(* CODESYS project stringhandler.library
   Company: KOSTAL GmbH & Co.KG
   Version: 2019.3.4.0
   DefaultNamespace: KOSTAL.TC3.Components.Stringhandler
   Title: KOSTAL.TC3.Components.Stringhandler
   Placeholder: KOSTAL.TC3.Components.Stringhandler
   Author: Frank Dümpelmann
   DocFormat: reStructuredText

Project tree, tasks and I/O mapping:
  libraries: KOSTAL.TC3.Components.listOfString, 2019.2.2.0 (KOSTAL GmbH & Co.KG); KOSTAL.TC3.Core.functionResponse, 2019.0.3.0 (KOSTAL GmbH & Co.KG); KOSTAL.TC3.Core.Settings, 2019.0.1.0 (KOSTAL GmbH & Co.KG); Tc2_Math, 3.3.1.0 (Beckhoff Automation GmbH); Tc2_Standard, 3.3.3.0 (Beckhoff Automation GmbH); Tc2_System, 3.4.26.0 (Beckhoff Automation GmbH); Tc2_Utilities, 3.3.54.0 (Beckhoff Automation GmbH); Tc3_Module, 3.3.21.0 (Beckhoff Automation GmbH)
  DUT/
    data type E_ALIGNMENT
  POU/
    obsolete/
      function F_CONCAT [ST]
      function F_Format [ST]
      function F_Text_Clear [ST]
      function block FB_Split [ST]: _pResult_clear, _settingsControl, Delimiter, pResults, sizeOfResultArray, split, status
    function F_FLOAT_TO_STRING [ST]
    function F_FormatMask [ST]
    function F_FormatNoMask [ST]
    function F_LCASE [ST]
    function F_LREAL_TO_STRING [ST]
    function F_REAL_TO_STRING [ST]
    function F_Replace [ST]
    function F_UCASE [ST]
    function block FB_CONCAT [ST]: addContent, clear, FB_exit, getResult, new
    function block FB_SplitEx [ST]: _settingsControl, clear, Delimiter, FB_exit, FB_init, getElement, maxElement, setElement, split, status
    function block FB_UrlEscape [ST]: Execute
  Project Information/
    function F_GetCompany [ST]
    function F_GetTitle [ST]
    function F_GetVersion [ST]
  Version/
    global variables Global_Version
  global variables GVL_CONSTANT
*)

// DUT/E_ALIGNMENT
TYPE E_ALIGNMENT :
	(
		LEFT 	:= 0,
		RIGHT	:= 1,
		CENTER	:= 2
	);
END_TYPE

// Version/Global_Version
{attribute 'TcGenerated'}
{attribute 'no-analysis'}
{attribute 'linkalways'}
// This function has been automatically generated from the project information.
VAR_GLOBAL CONSTANT
	{attribute 'const_non_replaced'}
	stLibVersion_KOSTAL_TC3_Components_Stringhandler : ST_LibVersion := (iMajor := 2019, iMinor := 3, iBuild := 4, iRevision := 0, nFlags := 1, sVersion := '2019.3.4.0');
END_VAR

// GVL_CONSTANT
{attribute 'qualified_only'}
VAR_GLOBAL CONSTANT
	
(*
65 A 	97 a 
66 B 	98 b 
67 C 	99 c 
68 D 	100 d 
69 E 	101 e 
70 F 	102 f 
71 G 	103 g 
72 H 	104 h 
73 I 	105 i 
74 J 	106 j 
75 K 	107 k 
76 L 	108 l 
77 M 	109 m 
78 N 	110 n 
79 O 	111 o 
80 P 	112 p 
81 Q 	113 q 
82 R 	114 r 
83 S 	115 s 
84 T 	116 t 
85 U 	117 u 
86 V 	118 v 
87 W 	119 w 
88 X 	120 x 
89 Y 	121 y 
90 Z 	122 z
*)

	START_UCASE	: BYTE:= 65;	//BYTE:= 65
	END_UCASE		: BYTE:= 90;	//BYTE:= 90
	START_LCASE	: BYTE:= 97;	//BYTE:= 97
	END_LCASE		: BYTE:= 122;	//BYTE:= 122
	OFFSET			: BYTE:= 32;	//BYTE:= 32

	OVERFLOW	: STRING:= 'OVERFLOW';
	
END_VAR

// POU/obsolete/F_CONCAT
(*

:Author: Frank Dümpelmann <f.duempelmann@kostal.com>, Martin Hundt <m.hundt@kostal.com>
:Date: 2018-10-29

Function
========
Concatination of variable number of lines to one line with maximum 255 chars

Usage notes
===============
Won't work with arrays shorter than 255 chars

Parameters
======================
| P_Line_1		: POINTER TO STRING(255) - Pointer to first element of an array[1..numberOfLines] OF STRING(255)
| numberOfLines	: USINT - defines the number of elements of the Array 

Return Value
============
String(255) - Concatination of the array's elements

Usage sample:
=============

.. code:: 

	PROGRAM MAIN
	VAR
		_aStrings	: ARRAY [0..4] OF STRING(255);
		_output 	: STRING(255); 
	END_VAR
	
	_aStrings[0] := 'Kostal';
	_aStrings[1] := ' ';
	_aStrings[2] := 'Automobil';
	_aStrings[3] := ' ';
	_aStrings[4] := 'Elektrik';
	
	_output := F_CONCAT(ADR(_aStrings[0]), 5);

*)

{attribute 'obsolete' := 'use instead FB_CONCAT'} 
FUNCTION F_CONCAT : KOSTAL_TC3_Core_Settings.T_MaxString

VAR_INPUT
	P_Line_1			: POINTER TO KOSTAL_TC3_Core_Settings.T_MaxString;	//Pointer to first Element  Array[1..numberOfLines] OF KOSTAL_TC3_Core_Settings.T_MaxString
	numberOfLines	: USINT;	// defines the number of Indices of the Array 
END_VAR

VAR
	_P_Line	: POINTER TO KOSTAL_TC3_Core_Settings.T_MaxString;
	_index	: UDINT;
END_VAR


F_CONCAT:= '';

IF P_Line_1 = 0 			THEN	RETURN;	END_IF
IF numberOfLines = 0 	THEN	RETURN;	END_IF


FOR _index:= 1 TO numberOfLines DO
	_P_line:= P_Line_1 + ((_index - 1) * SIZEOF(P_Line_1^));
	F_CONCAT:= CONCAT(F_CONCAT, _P_line^);
END_FOR

END_FUNCTION

// POU/FB_CONCAT
(*

:Author: Frank Dümpelmann <f.duempelmann@kostal.com>, Martin Hundt <m.hundt@kostal.com>
:Date: 2018-10-30

Function
========
| Function block to concatinate a variable number of strings
| Create a new array using the new method
| Add strings with addContent
| Receive the concatinated strings with getResult

Methods and Properties
======================
| See bottom of this document for a detailed description of each method or property

Usage sample:
=============

.. code:: 

	PROGRAM MAIN
	VAR
		_concat	: FB_CONCAT;
		_testConcat: STRING(255);
	END_VAR
	
	_concat.new(numberOfElements := 3);
	_concat.addContent(elementNumber := 1, text := '123');
	_concat.addContent(elementNumber := 2, text := '456');
	_concat.addContent(elementNumber := 3, text := '789');
	
	_testConcat := _concat.getResult();

*)

FUNCTION_BLOCK PUBLIC FB_CONCAT
VAR_INPUT
END_VAR
VAR_OUTPUT
END_VAR
VAR
	_pStack	: POINTER TO KOSTAL_TC3_Core_Settings.T_MaxString;
	_numberOfElements	: UINT;
END_VAR

(*
Description
===========
| Adds a string to the concatination stack at a certain position
| Existing content of the position will be overwritten
| Parameters:
| 	elementNumber : UINT - Position to insert the string (1-based)
| 	text : STRING(255) - String to insert
| Return value: BOOL - TRUE=String successfully added, FALSE=elementNumber invalid
*)

METHOD PUBLIC addContent : BOOL
VAR_INPUT
	elementNumber	: UINT;
	text					: KOSTAL_TC3_Core_Settings.T_MaxString;
END_VAR

IF _pStack = 0 THEN addContent:= FALSE;	RETURN;	END_IF

IF (elementNumber = 0) OR (elementNumber > _numberOfElements) THEN addContent:= FALSE;	RETURN;	END_IF

_pStack[elementNumber - 1]:= text;

addContent:= TRUE;
END_METHOD

(*
Description
===========
| Clear the concatination stack
*)

METHOD PUBLIC clear
VAR_INPUT
END_VAR

IF (_pStack <> 0) THEN	__DELETE(_pStack); END_IF
END_METHOD

(*
Description
===========
| Is called automatically
*)
METHOD FB_exit : BOOL
VAR_INPUT
	bInCopyCode : BOOL; // if TRUE, the exit method is called for exiting an instance that is copied afterwards (online change).
END_VAR

IF (_pStack <> 0) THEN __DELETE(_pStack);	END_IF
END_METHOD

(*
Description
===========
| Returns the concatinated strings
| Return value: STRING(255)
*)

METHOD PUBLIC getResult : KOSTAL_TC3_Core_Settings.T_MaxString
VAR_INPUT
END_VAR

VAR
	_i: UINT;
END_VAR

getResult:= '';	

IF _pStack = 0 THEN RETURN;	END_IF

FOR _i:= 0 TO _numberOfElements - 1 DO
	getResult:= CONCAT(getResult, _pStack[_i]);	
END_FOR
END_METHOD

(*
Description
===========
| Creates a new concatination stack
| Return value: BOOL -  FALSE=allocation has failed
*)

METHOD PUBLIC new: BOOL
VAR_INPUT
	numberOfElements	: UINT;
END_VAR


IF (_pStack <> 0) THEN __DELETE(_pStack);	END_IF

_numberOfElements:= numberOfElements;

IF _numberOfElements = 0 THEN
	_pStack:= 0;
ELSE
	_pStack:= __NEW(KOSTAL_TC3_Core_Settings.T_MaxString,_numberOfElements);
END_IF

new:= _pStack <> 0;
END_METHOD

END_FUNCTION_BLOCK

// POU/obsolete/F_Format
(*

:Author: Frank Dümpelmann <f.duempelmann@kostal.com>, Martin Hundt <m.hundt@kostal.com>
:Date: 2018-10-29

Function
========
| Formats =line= to the length of =mask= with the characters defined in =mask= and given =alignment=
| If =line= is longer than =mask=, the method will return =line= with the original length

Methods and Properties
======================
| line	: STRING(255) - String to format
| mask	: STRING(255) - e.g., '00000' formats line to 5 characters, filling up with the placeholder 0 
| alignment	: E_ALIGNMENT - Alignment of the original string

Usage sample:
=============

.. code:: 

	PROGRAM MAIN
	VAR	
		_Test : STRING(255) := 'test';
	END_VAR
	
	_Test := F_Format(line := _Test, mask:= 'xxxxxxxxxx', alignment:=E_ALIGNMENT.Left);

*)


{attribute 'obsolete' := 'Function was renamed to F_FormatMask'} 
FUNCTION F_Format : KOSTAL_TC3_Core_Settings.T_MaxString
VAR_INPUT
	line	: KOSTAL_TC3_Core_Settings.T_MaxString;	//
	mask	: KOSTAL_TC3_Core_Settings.T_MaxString;			//f.a. '00000' defines the minimum lenght and placeholder for empty string position 
	alignment	: E_ALIGNMENT;
END_VAR
VAR
END_VAR


F_Format:= F_FormatMask(line, mask, alignment);

(*
IF alignment = E_ALIGNMENT.LEFT THEN

	IF Tc2_Standard.LEN(mask) > Tc2_Standard.LEN(line) THEN
		F_Format:= Tc2_Standard.LEFT(Tc2_Standard.CONCAT(line, mask), Tc2_Standard.LEN(mask));		
	ELSE
		F_Format:= Tc2_Standard.LEFT(Tc2_Standard.CONCAT(line, mask), Tc2_Standard.LEN(line));		
	END_IF
	
ELSIF alignment = E_ALIGNMENT.RIGHT THEN

	IF Tc2_Standard.LEN(mask) > Tc2_Standard.LEN(line) THEN
		F_Format:= Tc2_Standard.RIGHT(Tc2_Standard.CONCAT(mask, line), Tc2_Standard.LEN(mask));		
	ELSE
		F_Format:= Tc2_Standard.RIGHT(Tc2_Standard.CONCAT(mask, line), Tc2_Standard.LEN(line));		
	END_IF

ELSE
	F_Format:= '';		
END_IF
*)

END_FUNCTION

// POU/F_FormatMask
(*

:Author: Frank Dümpelmann <f.duempelmann@kostal.com>, Martin Hundt <m.hundt@kostal.com>
:Date: 2018-10-29

Function
========
| Formats =line= to the length of =mask= with the characters defined in =mask= and given =alignment=
| If =line= is longer than =mask=, the method will return =line= with the original length

Methods and Properties
======================
| line	: STRING(255) - String to format
| mask	: STRING(255) - e.g., '00000' formats line to 5 characters, filling up with the placeholder 0 
| alignment	: E_ALIGNMENT - Alignment of the original string

Usage sample:
=============

.. code:: 

	PROGRAM MAIN
	VAR	
		_Test : STRING(255) := 'test';
	END_VAR
	
	_Test := F_Format(line := _Test, mask:= 'xxxxxxxxxx', alignment:=E_ALIGNMENT.Left);

*)


FUNCTION F_FormatMask : KOSTAL_TC3_Core_Settings.T_MaxString
VAR_INPUT
	line	: KOSTAL_TC3_Core_Settings.T_MaxString;	//
	mask	: KOSTAL_TC3_Core_Settings.T_MaxString;			//f.a. '00000' defines the minimum lenght and placeholder for empty string position 
	alignment	: E_ALIGNMENT;
END_VAR
VAR
END_VAR


IF alignment = E_ALIGNMENT.LEFT THEN

	IF Tc2_Standard.LEN(mask) > Tc2_Standard.LEN(line) THEN
		F_FormatMask:= Tc2_Standard.LEFT(Tc2_Standard.CONCAT(line, mask), Tc2_Standard.LEN(mask));		
	ELSE
		F_FormatMask:= Tc2_Standard.LEFT(Tc2_Standard.CONCAT(line, mask), Tc2_Standard.LEN(line));		
	END_IF
	
ELSIF alignment = E_ALIGNMENT.RIGHT THEN

	IF Tc2_Standard.LEN(mask) > Tc2_Standard.LEN(line) THEN
		F_FormatMask:= Tc2_Standard.RIGHT(Tc2_Standard.CONCAT(mask, line), Tc2_Standard.LEN(mask));		
	ELSE
		F_FormatMask:= Tc2_Standard.RIGHT(Tc2_Standard.CONCAT(mask, line), Tc2_Standard.LEN(line));		
	END_IF

ELSE
	F_FormatMask:= '';		
END_IF

END_FUNCTION

// POU/obsolete/F_Text_Clear
(*

:Author: Frank Dümpelmann <f.duempelmann@kostal.com>, Martin Hundt <m.hundt@kostal.com>
:Date: 2018-10-29

Function
========
Clear lines from an array of strings

Usage notes
===============
Won't work with arrays shorter than 255 chars

Parameters
======================
| P_Line_1		: POINTER TO STRING(255) - Pointer to first element of an array[1..numberOfLines] OF STRING(255)
| numberOfLines	: USINT - number of lines to clear 

Return Value
============
BOOL - TRUE=Array was cleared, FALSE=Pointer or array was empty

*)
{attribute 'obsolete' := 'Dangerous if wrong Pointer is set on P_Line_1'} 
FUNCTION F_Text_Clear : BOOL

VAR_INPUT
	P_Line_1			: POINTER TO KOSTAL_TC3_Core_Settings.T_MaxString;	//Pointer to first Element  Array[1..numberOfLines] OF STRING(255)
	numberOfLines	: USINT;	// defines the number of Indices of the Array 
END_VAR

VAR
	_P_Line	: POINTER TO KOSTAL_TC3_Core_Settings.T_MaxString;
	_index: UDINT;
END_VAR


F_Text_Clear:= FALSE;

IF P_Line_1 = 0 			THEN	RETURN;	END_IF
IF numberOfLines = 0 	THEN	RETURN;	END_IF

F_Text_Clear:= TRUE;

FOR _index:= 1 TO numberOfLines DO
	_P_line:= P_Line_1 + ((_index - 1) * SIZEOF(P_Line_1^) );
	_P_line^:= '';
END_FOR

END_FUNCTION

// POU/obsolete/FB_Split
(*

:Author: Frank Dümpelmann <f.duempelmann@kostal.com>, Martin Hundt <m.hundt@kostal.com>
:Date: 2018-10-30

Function
========
Function block to split a KOSTAL_TC3_Core_Settings.T_MaxString devided by a defined delimiter to an array of strings 

Usage notes
===============
| Create an array of String(255) for the results outside  FB_Split
| Set properties pResults and sizeOfResultArray
| Call Method split(in := string(255))
| If the result array is too small for the found elements, it is filled to its last element, 
| and an error message (status.success = false) is generated.

Methods and Properties
======================
| See bottom of this document for a detailed description of each method or property
| Methods starting with an underline(_) are internally used and can be ignored by the user

Usage sample:
=============

.. code:: 

	PROGRAM MAIN
	VAR
		_split : FB_Split;
		_splitString : STRING(255) := 'abc;def;ghi;jkl;mno;pqr;stu;vwx;yz';
		_splitArray : ARRAY[1..9] OF STRING(255);
	END_VAR
	
	_split.pResults := ADR(_splitArray[1]);
	_split.sizeOfResultArray := 10;
	_split.split(in:=_splitString);

*)
{attribute 'obsolete' := 'use instead FB_SplitEx'} 
FUNCTION_BLOCK PUBLIC FB_Split

VAR
	
	_Delimiter	: STRING(1):= ';';	//STRING(1):= ';'
	_pResults	: POINTER TO KOSTAL_TC3_Core_Settings.T_MaxString;	//>> Pointer to first Element of Array OF KOSTAL_TC3_Core_Settings.T_MaxString
	_sizeOfResultArray	: UINT;	//UINT	>>	size of result Array OF String(255)

	_IN	: KOSTAL_TC3_Core_Settings.T_MaxString;

	_status	: KOSTAL_TC3_Core_functionResponse.FB_functionResponse;	//KOSTAL_functionResponse.FB_functionResponse

END_VAR

METHOD PROTECTED _pResult_clear
VAR_INPUT
END_VAR

VAR
	_index: INT;	//INT
	_pResultsToClear	: POINTER TO KOSTAL_TC3_Core_Settings.T_MaxString;
END_VAR

_pResultsToClear:= _pResults;

FOR _index:= 0 TO UINT_TO_INT(_sizeOfResultArray - 1) DO
	_pResultsToClear	:= _pResults + INT_TO_DWORD(_index * 256);
	_pResultsToClear^	:= '';
END_FOR
END_METHOD

METHOD PROTECTED _settingsControl : KOSTAL_TC3_Core_functionResponse.FB_functionResponse
VAR_INPUT
END_VAR


IF _pResults = 0 THEN
	_settingsControl.status	:= 'Pointer >pResults< is invalid';
	_settingsControl.success:= FALSE;
	RETURN;
END_IF

IF _sizeOfResultArray <= 0 THEN
	_settingsControl.status	:= '>sizeOfResultArray< is invalid';
	_settingsControl.success:= FALSE;
	RETURN;
END_IF

IF _Delimiter = '' THEN
	_settingsControl.status	:= '>Delimiter< is invalid';
	_settingsControl.success:= FALSE;
	RETURN;
END_IF

_settingsControl.status	:= '';
_settingsControl.success:= TRUE;
END_METHOD

(*
Description
===========
| Delimiter deviding the elements in the string
| Attention: Only ONE character!
| default: ';'
*)

PROPERTY PUBLIC Delimiter : STRING(1)
GET

Delimiter:= _Delimiter;
END_GET
SET

_Delimiter:= Delimiter;
END_SET
END_PROPERTY

(*
Description
===========
| Pointer to Array of String(255)
| Pointer to the first element of the results array
*)
PROPERTY PUBLIC pResults : POINTER TO KOSTAL_TC3_Core_Settings.T_MaxString
GET

pResults:= _pResults;
END_GET
SET

_pResults:= pResults;
END_SET
END_PROPERTY

(*
Description
===========
| Number of elements in pResults 
*)
PROPERTY PUBLIC sizeOfResultArray : UINT
GET

sizeOfResultArray:= _sizeOfResultArray;
END_GET
SET

_sizeOfResultArray:= sizeOfResultArray;
END_SET
END_PROPERTY

(*
Description
===========
| Splits the string to the array
*)

METHOD PUBLIC split 

VAR_INPUT
	IN	: KOSTAL_TC3_Core_Settings.T_MaxString;
END_VAR

VAR
	_resultIndex	: UINT;
	_signCount		: UINT;
	
	_pIN_BYTE		: POINTER TO BYTE;

	_pOne_CHAR							: POINTER TO BYTE;
	_pOne_CHAR_Termination	: POINTER TO BYTE;
	_One_CHAR								: STRING(1);

	_IN_Count		: UINT;
	
	_pResultElement	: POINTER TO KOSTAL_TC3_Core_Settings.T_MaxString;
END_VAR

_status:= _settingsControl();

IF NOT _status.success THEN RETURN;	END_IF

_pResult_clear();

IF IN = '' THEN
	_status.status	:= '>IN< is empty';
	_status.success:= TRUE;
	RETURN;
END_IF

_pIN_BYTE	:= ADR(IN);
_One_CHAR:= '';
_pOne_CHAR	:= ADR(_One_CHAR);
_pOne_CHAR_Termination:= _pOne_CHAR + 1;

_resultIndex		:= 0;
_signCount:= 0;


FOR _IN_Count:= 0 TO INT_TO_UINT(LEN(IN)) - 1 DO


	IF _resultIndex > (_sizeOfResultArray - 1) THEN
		_status.status	:= '>IN< contains to much elements';
		_status.success:= FALSE;
		RETURN;
	END_IF

	
	_pIN_BYTE		:= ADR(IN) + UINT_TO_DWORD(_IN_Count);
	_pOne_CHAR^	:= _pIN_BYTE^;
	_pOne_CHAR_Termination^	:= 0;
	
	_pResultElement:= _pResults + UINT_TO_DWORD(_resultIndex * SIZEOF(IN));

	IF _pIN_BYTE^ = 0 THEN
		_status.status	:= 'end of line reached';
		_status.success:= TRUE;
		RETURN;
	END_IF
	
	
	IF _One_CHAR = _Delimiter THEN

		_resultIndex:= _resultIndex + 1;
		
	ELSE
		
		_pResultElement^:=	CONCAT(_pResultElement^, _One_CHAR);
		
	END_IF
	
	
END_FOR

_status.status	:= CONCAT(UINT_TO_STRING(_resultIndex + 1), ' Element(s) found');
_status.success	:= TRUE;
END_METHOD

(*
Description
===========
| Success: BOOL - Split succeeded
| Status: 
| Success = TRUE: Number of elements found
| Success = FALSE: Reason for failure
*)
PROPERTY PUBLIC status : REFERENCE TO KOSTAL_TC3_Core_functionResponse.FB_functionResponse
GET


status	REF= _status;
END_GET
END_PROPERTY

END_FUNCTION_BLOCK

// POU/FB_SplitEx
(*

:Author: Frank Dümpelmann <f.duempelmann@kostal.com>, Martin Hundt <m.hundt@kostal.com>
:Date: 2018-10-30

Function
========
Function block to split a KOSTAL_TC3_Core_Settings.T_MaxString devided by a defined delimiter to an ListOf Object 

Usage notes
===============
| Call Method split(in := string(255))

Methods and Properties
======================
| See bottom of this document for a detailed description of each method or property
| Methods starting with an underline(_) are internally used and can be ignored by the user

Usage sample:
=============

.. code:: 

	PROGRAM MAIN
	VAR
		_split : FB_Split;
		_splitString : KOSTAL_TC3_Core_Settings.T_MaxString := 'abc;def;ghi;jkl;mno;pqr;stu;vwx;yz';
	END_VAR
	
	_split.split(in:=_splitString);

*)
FUNCTION_BLOCK PUBLIC FB_SplitEx

VAR
	
	_Delimiter	: STRING(1):= ';';	//STRING(1):= ';'

	_IN	: KOSTAL_TC3_Core_Settings.T_MaxString;

	_status			: KOSTAL_TC3_Core_functionResponse.FB_functionResponse;

	_results		: KOSTAL_TC3_Components_listOfString.FB_ListOfString_255;
	_maxElement	: UINT;
	
END_VAR

METHOD PROTECTED _settingsControl : KOSTAL_TC3_Core_functionResponse.FB_functionResponse
VAR_INPUT
END_VAR


IF _Delimiter = '' THEN
	_settingsControl.status	:= '>Delimiter< is invalid';
	_settingsControl.success:= FALSE;
	RETURN;
END_IF

IF _Delimiter = '' THEN
	_status.status	:= '>Delimiter< is invalid';
	_status.success:= FALSE;
	RETURN;
END_IF

_settingsControl.status	:= '';
_settingsControl.success:= TRUE;
END_METHOD

METHOD PUBLIC clear
VAR_INPUT
END_VAR

_results.clear();
END_METHOD

(*
Description
===========
| Delimiter deviding the elements in the string
| Attention: Only ONE character!
| default: ';'
*)

PROPERTY PUBLIC Delimiter : STRING(1)
GET

Delimiter:= _Delimiter;
END_GET
SET

_Delimiter:= Delimiter;
END_SET
END_PROPERTY

METHOD FB_exit : BOOL
VAR_INPUT
	bInCopyCode : BOOL; // if TRUE, the exit method is called for exiting an instance that is copied afterwards (online change).
END_VAR

_results.clear();
END_METHOD

METHOD FB_init : BOOL
VAR_INPUT
	bInitRetains : BOOL; // if TRUE, the retain variables are initialized (warm start / cold start)
	bInCopyCode : BOOL;  // if TRUE, the instance afterwards gets moved into the copy code (online change)
END_VAR

_results.clear();
END_METHOD

METHOD PUBLIC getElement : KOSTAL_TC3_Core_Settings.T_MaxString
VAR_INPUT
	elementNumber	: UINT;
END_VAR

IF (elementNumber = 0) OR (elementNumber > _results.numberOfLines_GET()) THEN
	getElement:= '';
ELSE
	getElement:= _results.line_GET(numberOfLine:= elementNumber);
END_IF
END_METHOD

METHOD PUBLIC maxElement : UINT
VAR_INPUT
END_VAR

maxElement:= _results.numberOfLines_GET();
END_METHOD

METHOD PUBLIC setElement : BOOL
VAR_INPUT
	line	: KOSTAL_TC3_Core_Settings.T_MaxString;
	elementNumber	: UINT;
END_VAR

IF (elementNumber = 0) OR (elementNumber > _results.numberOfLines_GET()) THEN
	setElement:= FALSE;
ELSE
	_results.line_SET(line:= line, numberOfLine:= elementNumber);
	setElement:= TRUE; 
END_IF
END_METHOD

(*
Description
===========
| Splits the string to the array
*)

METHOD PUBLIC split 

VAR_INPUT
	IN	: KOSTAL_TC3_Core_Settings.T_MaxString;
END_VAR

VAR
	_delimiterPosition: INT;
END_VAR

_status:= _settingsControl();

IF NOT _status.success THEN RETURN;	END_IF

_results.clear();

IF IN = '' THEN
	_status.status	:= '>IN< is empty';
	_status.success:= TRUE;
	RETURN;
END_IF

_IN:= IN;


REPEAT

	_delimiterPosition:= FIND(STR1:= _IN, STR2:= _Delimiter);

	IF _delimiterPosition = 0 THEN
 		_results.addLine(_IN);
	ELSE
 		_results.addLine(newLine:= Tc2_Standard.LEFT(_IN, _delimiterPosition - 1));
		_IN:= Tc2_Standard.RIGHT(STR:= _IN, SIZE:= Tc2_Standard.LEN(_IN) - _delimiterPosition);
	END_IF
		
UNTIL	_delimiterPosition = 0
END_REPEAT

_status.status	:= CONCAT(UINT_TO_STRING(_results.numberOfLines_GET()), ' Element(s) found');
_status.success	:= TRUE;
END_METHOD

(*
Description
===========
| Success: BOOL - Split succeeded
| Status: 
| Success = TRUE: Number of elements found
| Success = FALSE: Reason for failure
*)
PROPERTY PUBLIC status : REFERENCE TO KOSTAL_TC3_Core_functionResponse.FB_functionResponse
GET


status	REF= _status;
END_GET
END_PROPERTY

END_FUNCTION_BLOCK

// POU/F_FLOAT_TO_STRING
(*
Supported Data Types:
REAL;LREAL
*)

FUNCTION F_FLOAT_TO_STRING : STRING(512)

VAR_INPUT
	IN			: Tc2_Utilities.FLOAT;
	Digits	: INT;	//Number of digits after the decimal point
END_VAR

VAR
	(*
	_s					: STRING;
	_DINT				: DINT;
	_DINTdigits	: DINT;
	*)
	//_T_Arg: Tc2_Utilities.T_Arg;
	_IN			: LREAL;
END_VAR


_IN:= IN;

//_T_Arg:= Tc2_Utilities.F_LREAL(IN);

IF NOT Tc2_Utilities.LrealIsFinite(_IN) THEN	
	F_FLOAT_TO_STRING:= GVL_CONSTANT.OVERFLOW;
	RETURN;	
ELSIF Tc2_Utilities.LrealIsNaN(_IN) THEN	
	F_FLOAT_TO_STRING:= GVL_CONSTANT.OVERFLOW;
	RETURN;	
END_IF

F_FLOAT_TO_STRING:=Tc2_Utilities.LREAL_TO_FMTSTR(IN, Digits, FALSE);

(*
_s:='';

//Is in DINT Range?
IF (IN < REAL#-2147483648.0) 
OR (IN > REAL#2147483647.0)
OR (NOT Tc2_Utilities.IsFinite(Tc2_Utilities.F_LREAL(IN))) 
THEN 

	_s:= GVL_CONSTANT.OVERFLOW;
	
ELSE
	 
	_DINT				:= TRUNC(IN);
	_DINTdigits	:= LREAL_TO_DINT(ABS(Tc2_Math.FRAC(IN)) * EXPT(10, Digits));
	
	_s:= DINT_TO_STRING(_DINT);
	
	if Digits > 0 then
		_s:= Tc2_Standard.CONCAT(_s, '.');
		_s:= Tc2_Standard.CONCAT(_s, DINT_TO_STRING(_DINTdigits));
	END_IF

END_IF
*)

END_FUNCTION

// POU/F_FormatNoMask
(*

:Author: Martin Hundt <m.hundt@kostal.com>
:Date: 2021-12-10

Function
========
| Formats =line= to the length of =formatLength= with the characters =char= and given =alignment=
| If =line= is longer than =formatLength=, the method will return =line= with the original length

Methods and Properties
======================
| line			: STRING(255) - String to format
| formatLength	: UINT - length of formatted string 
| char			: STRING(1) - Character to fill the sting. Default: Space 
| alignment		: E_ALIGNMENT - Alignment of the return string

Usage sample:
=============
See best practice
*)


FUNCTION F_FormatNoMask : KOSTAL_TC3_Core_Settings.T_MaxString
VAR_INPUT
	line			: KOSTAL_TC3_Core_Settings.T_MaxString;	//
	formatLength	: UINT;
	char			: STRING(1); 
	alignment		: E_ALIGNMENT;
END_VAR
VAR
	_stringLength	: UINT;
	_fillLength		: UINT;
	_out			: KOSTAL_TC3_Core_Settings.T_MaxString;
	_i				: UINT;
END_VAR


IF char = '' THEN 
	char := ' '; 
END_IF
_stringLength := INT_TO_UINT(Tc2_Standard.LEN(line));

IF _stringLength >= formatLength THEN
	_out := line;
ELSIF alignment = E_ALIGNMENT.LEFT THEN
	_out := line;
	FOR _i:= _stringLength TO formatLength DO
		_out := Tc2_Standard.CONCAT(_out, char);
	END_FOR

	
ELSIF alignment = E_ALIGNMENT.RIGHT THEN
	
	FOR _i:= 1 TO (formatLength - _stringLength) DO
		_out := Tc2_Standard.CONCAT(_out, char);
	END_FOR
	_out := Tc2_Standard.CONCAT(_out, line);
	
ELSIF alignment = E_ALIGNMENT.CENTER THEN	
	
	_fillLength := (formatLength-_stringLength)/2;
	
	FOR _i:=0 TO formatLength DO	//Fill with spaces
		_out := CONCAT(_out, char);
	END_FOR
	
	
	_out :=  Tc2_Standard.INSERT(_out, line,_fillLength + 1);
		
END_IF

F_FormatNoMask:= _out;

END_FUNCTION

// POU/F_LCASE
(*

:Author: Frank Dümpelmann <f.duempelmann@kostal.com>, Martin Hundt <m.hundt@kostal.com>
:Date: 2018-10-30

Function
========
Set all characters in the string to lower case

Usage notes
===============
| Only ASCII charset is supported

*) 
FUNCTION F_LCASE : KOSTAL_TC3_Core_Settings.T_MaxString
VAR_INPUT
	IN		: KOSTAL_TC3_Core_Settings.T_MaxString;
END_VAR

VAR
	_pos	: INT;
	_sign	: STRING(1);
END_VAR


IF IN <> '' THEN

	FOR _pos:= 1 TO LEN(IN) DO
		_sign:= MID(IN,1,_pos);
		IF F_ToASC(_sign) >= GVL_CONSTANT.START_UCASE AND F_ToASC(_sign) <= GVL_CONSTANT.END_UCASE THEN
			_sign:= F_ToCHR(F_ToASC(_sign) + GVL_CONSTANT.OFFSET);
			IN:= REPLACE(IN, _sign, 1, _pos);
		END_IF;
	END_FOR;

END_IF;

F_LCASE:= IN;

END_FUNCTION

// POU/F_LREAL_TO_STRING
(*
Supported Data Types:
REAL;LREAL
*)

FUNCTION F_LREAL_TO_STRING : STRING(512)

VAR_INPUT
	IN			: LREAL;
	Digits	: INT;	//Number of digits after the decimal point
END_VAR

VAR
	(*
	_s					: STRING;
	_DINT				: DINT;
	_DINTdigits	: DINT;
	*)
	//_T_Arg: Tc2_Utilities.T_Arg;
	_IN			: LREAL;
END_VAR


_IN:= IN;

//_T_Arg:= Tc2_Utilities.F_LREAL(IN);

IF NOT Tc2_Utilities.LrealIsFinite(_IN) THEN	
	F_LREAL_TO_STRING:= GVL_CONSTANT.OVERFLOW;
	RETURN;	
ELSIF Tc2_Utilities.LrealIsNaN(_IN) THEN	
	F_LREAL_TO_STRING:= GVL_CONSTANT.OVERFLOW;
	RETURN;	
END_IF

F_LREAL_TO_STRING:=Tc2_Utilities.LREAL_TO_FMTSTR(IN, Digits, FALSE);

(*
_s:='';

//Is in DINT Range?
IF (IN < REAL#-2147483648.0) 
OR (IN > REAL#2147483647.0)
OR (NOT Tc2_Utilities.IsFinite(Tc2_Utilities.F_LREAL(IN))) 
THEN 

	_s:= GVL_CONSTANT.OVERFLOW;
	
ELSE
	 
	_DINT				:= TRUNC(IN);
	_DINTdigits	:= LREAL_TO_DINT(ABS(Tc2_Math.FRAC(IN)) * EXPT(10, Digits));
	
	_s:= DINT_TO_STRING(_DINT);
	
	if Digits > 0 then
		_s:= Tc2_Standard.CONCAT(_s, '.');
		_s:= Tc2_Standard.CONCAT(_s, DINT_TO_STRING(_DINTdigits));
	END_IF

END_IF
*)

END_FUNCTION

// POU/F_REAL_TO_STRING
(*
Supported Data Types:
REAL;LREAL
*)
FUNCTION F_REAL_TO_STRING : STRING(512)

VAR_INPUT
	IN			: REAL;
	Digits	: INT;	//Number of digits after the decimal point
END_VAR

VAR
	(*
	_s					: STRING;
	_DINT				: DINT;
	_DINTdigits	: DINT;
	*)
	_T_Arg: Tc2_Utilities.T_Arg;
END_VAR




_T_Arg:= Tc2_Utilities.F_REAL(IN);

IF NOT Tc2_Utilities.IsFinite(_T_Arg) THEN	
	F_REAL_TO_STRING:= GVL_CONSTANT.OVERFLOW;
	RETURN;	
END_IF

F_REAL_TO_STRING:=Tc2_Utilities.LREAL_TO_FMTSTR(IN, Digits, FALSE);


(*
_s:='';

//Is in DINT Range?

//IF (IN < REAL#-2147483648.0) 
//OR (IN > REAL#2147483647.0) 

IF 		(NOT Tc2_Utilities.IsFinite(Tc2_Utilities.F_REAL(IN)))								THEN	_s:= GVL_CONSTANT.OVERFLOW;  
ELSIF (NOT Tc2_Utilities.IsFinite(Tc2_Utilities.F_DINT(REAL_TO_DINT(IN))))	THEN	_s:= GVL_CONSTANT.OVERFLOW; 
ELSE
	
	_DINT				:= TRUNC(IN);
	_DINTdigits	:= REAL_TO_DINT(ABS(Tc2_Math.FRAC(IN)) * EXPT(10, Digits));
	
	_s:= DINT_TO_STRING(_DINT);
	
	if Digits > 0 then
		_s:= Tc2_Standard.CONCAT(_s, '.');
		_s:= Tc2_Standard.CONCAT(_s, DINT_TO_STRING(_DINTdigits));
	END_IF
	
END_IF
*)

END_FUNCTION

// POU/F_Replace
(*

:Author: Frank Dümpelmann <f.duempelmann@kostal.com>, Martin Hundt <m.hundt@kostal.com>
:Date: 2018-10-30

Function
========
Replace all occurencies of a given string with another string

Methods and Properties
======================
| source 						: KOSTAL_TC3_Core_Settings.T_MaxString - string to replace in
| toReplace					: KOSTAL_TC3_Core_Settings.T_MaxString - string to replace
| replaceWith 			: KOSTAL_TC3_Core_Settings.T_MaxString - string to replace with
| numberOfReplaces	: Replace only the first X occurencies from left (default: -1, replace all occurrencies)

Usage sample:
=============

.. code:: 

	PROGRAM MAIN
	VAR	
		_replaceTest : KOSTAL_TC3_Core_Settings.T_MaxString;
	END_VAR
	
	_replaceTest := 'abcdefabcdefabcdef';
	_replaceTest := F_Replace(source := _replaceTest, toReplace := 'abc', replaceWith := 'xyz', numberOfReplaces := 1);
	;

*) 

FUNCTION F_Replace : KOSTAL_TC3_Core_Settings.T_MaxString

VAR_INPUT
	source						: KOSTAL_TC3_Core_Settings.T_MaxString;
	toReplace					: KOSTAL_TC3_Core_Settings.T_MaxString;
	replaceWith				: KOSTAL_TC3_Core_Settings.T_MaxString;
	numberOfReplaces	: INT:= -1;	(*INT:= -1 defines to replace all occurrences *)
END_VAR

VAR
	_index				: INT;
	_pos					: INT;
	_replaced			: KOSTAL_TC3_Core_Settings.T_MaxString;
	_toReplaceLen	: INT;
	_searchPos		: INT;
	_searchString	: KOSTAL_TC3_Core_Settings.T_MaxString;
	_i: INT;
END_VAR



IF 		numberOfReplaces  =  0  									THEN	F_Replace:= source;	RETURN;	//no replacement required
ELSIF Tc2_Standard.FIND(source, toReplace) = 0	THEN 	F_Replace:= source;	RETURN;	//no replacement required
ELSIF numberOfReplaces  <  0  									THEN	_index:= LEN(source);				//full replacement required
ELSE																									_index:= numberOfReplaces;	//replacement limmitted by numberOfReplaces
END_IF

//prepare
_replaced			:= '';
_toReplaceLen	:= Tc2_Standard.LEN(toReplace);
_searchString	:= source;
_searchPos		:= 1;


FOR _i:= 1 TO _index DO
	
	//find next to replace content
	_pos:= Tc2_Standard.FIND(_searchString, toReplace);

	//no further to replace found
	IF _pos = 0 THEN	EXIT;	END_IF
		
	//get left n characters until _pos
	IF _pos > 1 THEN	_replaced:= Tc2_Standard.CONCAT(_replaced, Tc2_Standard.LEFT(_searchString, _pos - 1));	END_IF

	//add replaced content
	_replaced:= Tc2_Standard.CONCAT(_replaced, replaceWith);
	
	//Capture the remaining characters to be checked   
	_searchString:= Tc2_Standard.RIGHT(_searchString, Tc2_Standard.LEN(_searchString) - (_pos - 1) - _toReplaceLen);
	
END_FOR

_replaced:= Tc2_Standard.CONCAT(_replaced, _searchString);
 	
F_Replace:= _replaced;

END_FUNCTION

// POU/F_UCASE
(*

:Author: Frank Dümpelmann <f.duempelmann@kostal.com>, Martin Hundt <m.hundt@kostal.com>
:Date: 2018-10-30

Function
========
Set all characters in the string to upper case

Usage notes
===============
| Only ASCII charset is supported

*) 

FUNCTION F_UCASE : KOSTAL_TC3_Core_Settings.T_MaxString

VAR_INPUT
	IN		: KOSTAL_TC3_Core_Settings.T_MaxString;
END_VAR

VAR
	_pos		: INT;
	_sign	: STRING(1);
END_VAR


IF IN <> '' THEN

	FOR _pos:= 1 TO LEN(IN) DO
		_sign:= MID(IN, 1, _pos);
		IF F_ToASC(_sign) >= GVL_CONSTANT.START_LCASE AND F_ToASC(_sign) <= GVL_CONSTANT.END_LCASE THEN
			_sign:= F_ToCHR(f_ToASC(_sign) - GVL_CONSTANT.OFFSET);
			IN:= REPLACE(IN, _sign, 1, _pos);
		END_IF;
	END_FOR;

END_IF;

F_UCASE:= IN;

END_FUNCTION

// POU/FB_UrlEscape
(*

:Author: Frank Dümpelmann <f.duempelmann@kostal.com>
:Date: 2018-10-30

Function
========
Class for replacing invalid characters in a URL with escape sequences. 
*)

FUNCTION_BLOCK PUBLIC FB_UrlEscape

VAR
	_s	: KOSTAL_TC3_Core_Settings.T_MaxString;
END_VAR

(*
Return TRUE 	: At least one character was escaped.
Return FALSE	: No character was escaped.
*)
METHOD PUBLIC Execute : BOOL

VAR_INPUT
	URL					: KOSTAL_TC3_Core_Settings.T_MaxString;
	URL_Escaped	: REFERENCE TO KOSTAL_TC3_Core_Settings.T_MaxString;	//Reference to a resultstring
END_VAR


//$24 (Hex) is ASCII Code for %

_s:= URL;

IF _s <> '' THEN

	_s:= F_Replace(_s,'%', '%25', -1);	
	
	_s:= F_Replace(_s,' ', '%20', -1);
	_s:= F_Replace(_s,'<', '%3C', -1);
	_s:= F_Replace(_s,'>', '%3E', -1);
	_s:= F_Replace(_s,'#', '%23', -1);
	_s:= F_Replace(_s,'+', '%2B', -1);
	_s:= F_Replace(_s,'{', '%7B', -1);
	_s:= F_Replace(_s,'}', '%7D', -1);
	_s:= F_Replace(_s,'|', '%7C', -1);
	_s:= F_Replace(_s,'\', '%5C', -1);
	_s:= F_Replace(_s,'^', '%5E', -1);
	_s:= F_Replace(_s,'~', '%7E', -1);
	_s:= F_Replace(_s,'[', '%5B', -1);
	_s:= F_Replace(_s,']', '%5D', -1);
	_s:= F_Replace(_s,'$'', '%60', -1);
	_s:= F_Replace(_s,';', '%3B', -1);
	_s:= F_Replace(_s,'/', '%2F', -1);
	_s:= F_Replace(_s,'?', '%3F', -1);
	_s:= F_Replace(_s,':', '%3A', -1);
	_s:= F_Replace(_s,'@', '%40', -1);
	_s:= F_Replace(_s,'=', '%3D', -1);
	_s:= F_Replace(_s,'&', '%26', -1);
	_s:= F_Replace(_s,'$$', '%24', -1);

END_IF

Execute:= _s <> URL;

IF __ISVALIDREF(URL_Escaped) THEN	URL_Escaped:= _s;	END_IF
END_METHOD

END_FUNCTION_BLOCK

// Project Information/F_GetCompany
// This function has been automatically generated from the project information.
{attribute 'signature_flag' := '1073741824'}
{attribute 'TcGenerated'}
{attribute 'no-analysis'}
FUNCTION F_GetCompany : WSTRING
VAR_INPUT
	
END_VAR

F_GetCompany := "KOSTAL GmbH & Co.KG";

END_FUNCTION

// Project Information/F_GetTitle
// This function has been automatically generated from the project information.
{attribute 'signature_flag' := '1073741824'}
{attribute 'TcGenerated'}
{attribute 'no-analysis'}
FUNCTION F_GetTitle : WSTRING
VAR_INPUT
	
END_VAR

F_GetTitle := "KOSTAL.TC3.Components.Stringhandler";

END_FUNCTION

// Project Information/F_GetVersion
// This function has been automatically generated from the project information.
{attribute 'signature_flag' := '1073741824'}
{attribute 'TcGenerated'}
{attribute 'no-analysis'}
FUNCTION F_GetVersion : ST_LibVersion
VAR_INPUT
	
END_VAR

F_GetVersion.iMajor := 2019;
F_GetVersion.iMinor := 3;
F_GetVersion.iBuild := 4;
F_GetVersion.iRevision := 0;
F_GetVersion.sVersion := '2019.3.4.0';
F_GetVersion.nFlags := 1;

END_FUNCTION
